FUNCTION_BLOCK T_SafeRTrig_UserFB EXTENDS T_SafeFunctionBlockBase
VAR_INPUT
	Signal : BOOL;
END_VAR
VAR_OUTPUT
	Trigger : BOOL;
END_VAR
VAR
	safeRs : T_SafeRs(_group);
	safeAnd : T_SafeAnd(_group);
END_VAR

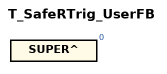
SUPER^();

METHOD FB_init : BOOL
VAR_INPUT
	bInitRetains	: BOOL;
	bInCopyCode	: BOOL;
	group	: REFERENCE TO T_SafeGroup;
END_VAR
safeRs.SetGroupReference(bInCopyCode := bInCopyCode, group := group);
safeAnd.SetGroupReference(bInCopyCode := bInCopyCode, group := group);
END_METHOD

METHOD PROTECTED Process
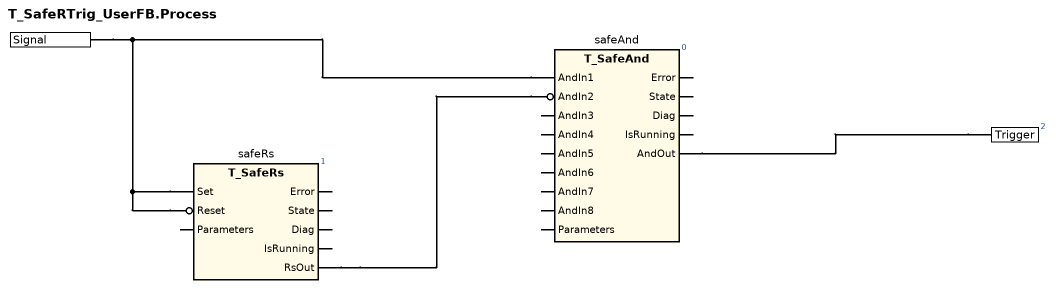
safeAnd(AndIn1 := Signal, AndIn2 := NOT safeRs.RsOut); // T_SafeAnd
safeRs(Set := Signal, Reset := NOT Signal); // T_SafeRs
Trigger := safeAnd.AndOut;
END_METHOD

END_FUNCTION_BLOCK

(* stored: Version 1.1.0.1
   POU T_SafeRTrig_UserFB: Id {9393d438-798f-49c8-973e-7f1078c0fc88}, SpecialFunc None
   Method FB_init: Id {d130f029-eff5-470e-9b9a-b39e1ab5c187}
   Method Process: Id {ee92d2ee-e173-411f-86da-1ebd8d2ff0c4} *)
